// TIA Portal V21 export
Screen "R03_BtnSet"  1024x768, Number=42, Template=Tpl
  ScreenLayer 
    Button "P_Btn" at 10,10 size 100x30  TextOff="BTN", TextOn="BTN"
      on Press: SetBit(Tag := P_SwOn)
